(* IEC 61131-3 sources: IRIS-Project/LASAL CONTROL SOFTWARE/LasalProject_2025_09_12/Runtime/%LASALAPPDATA%/Runtime/Library/Loader/Network, 1 file *)

(* ---- ConfigObjects.st ---- *)
FUNCTION GLOBAL TAB TASK_CONF
_K_TASK, _K_REAL,
_K_END_VAR,

_K_TASK, _K_CYCLIC,
_K_END_VAR,

_K_TASK, _K_BACKGROUND,
_K_END_VAR,

_K_END_CONF
END_FUNCTION

FUNCTION GLOBAL TAB IPR_CONF
_K_IPR
	0$UINT,
_K_END_VAR,
_K_END_CONF
END_FUNCTION

FUNCTION GLOBAL TAB CONFIG_TABLES
00033$UINT,
0$UINT, 1, 0, "_MULTITASK",
0$UINT, 1, 0, "_TASKOBJECTCONTROL",
0$UINT, 0, 0, "BASEIP",
0$UINT, 0, 0, "CLASSREADER",
0$UINT, 0, 0, "CONNECTREADER",
0$UINT, 1, 2, "DATASERVICE",
0$UINT, 0, 1, "DEBUGIP",
0$UINT, 0, 0, "INITREADER",
0$UINT, 0, 0, "IPRMGR",
0$UINT, 0, 0, "IPRREADER",
0$UINT, 1, 20, "MERKEREX",
0$UINT, 0, 0, "MMBUFFER",
0$UINT, 0, 0, "MMCONNECTIONHANDLER",
0$UINT, 0, 0, "MMCONNECTIONREADER",
0$UINT, 0, 0, "MMSERVER",
0$UINT, 0, 0, "MMSERVER4BYTEIMPL",
0$UINT, 0, 0, "MMSERVERIMPL",
0$UINT, 0, 0, "MMSERVERMERKEREX",
0$UINT, 0, 0, "MMSERVERREADER",
0$UINT, 0, 0, "MMSERVERSTRING",
0$UINT, 0, 0, "MMSTATION",
0$UINT, 0, 0, "MMSTATIONREADER",
0$UINT, 0, 1, "OBJECTREADER",
0$UINT, 0, 0, "PROGIP",
0$UINT, 0, 0, "PROGMGR",
0$UINT, 0, 0, "PROJECTREADER",
0$UINT, 0, 0, "PTRCHK",
0$UINT, 1, 16, "RAMEX",
0$UINT, 0, 1, "RETSVRFILE",
0$UINT, 1, 1, "RETSVRRAM",
0$UINT, 1, 82, "STRINGINTERNAL",
0$UINT, 0, 0, "TASKREADER",
0$UINT, 1, 3, "VIRTUALBASEINIT",
TASK_CFG$UINT, 0, 0, "TASK_CONF",
IPR_CFG$UINT, 0, 0, "IPR_CONF",
PRJ_CFG$UINT, 0, 0, "Loader",
END_FUNCTION
